(* IEC 61131-3 sources: plcassist-cli/packages/volt-lsp-iec/test-corpus/lenze-mid/Device/Plc Logic/Application/Library Manager/(unresolved)/visuusermgmt3 interfaces, 17 files *)

(* ---- VUM_CONSTANTS.gvl ---- *)
VAR_GLOBAL
	VISU_VUM_MAX_GROUPS_PER_USER : INT := 10;
END_VAR

(* ---- IEXTERNALUSERDATABASEPROVIDER.itf ---- *)
INTERFACE IEXTERNALUSERDATABASEPROVIDER
END_INTERFACE

METHOD CHANGEUSERPASSWORD : VUM_ReturnValues
VAR_INPUT
	WSTUSERNAME : WSTRING;
	WSTNEWPASSWORD : WSTRING;
	WSTOLDPASSWORD : WSTRING;
END_VAR
END_METHOD

METHOD CHECKLOGIN : VUM_ReturnValues
VAR_INPUT
	WSTUSERNAME : WSTRING;
	WSTPASSWORD : WSTRING;
END_VAR
VAR_OUTPUT
	WSTFULLNAME : WSTRING;
	DWUSERGROUPID : DWORD;
END_VAR
END_METHOD

METHOD CHECKLOGINWITHGROUPID : VUM_ReturnValues
VAR_INPUT
	WSTUSERNAME : WSTRING;
	WSTPASSWORD : WSTRING;
	DWUSERGROUPID : DWORD;
END_VAR
VAR_OUTPUT
	WSTFULLNAME : WSTRING;
END_VAR
END_METHOD

METHOD CHANGEUSER : VUM_ReturnValues
VAR_INPUT
	PVUMUSER : POINTER TO VUM_User;
	UDIINDEX : UDINT;
	EEDITTYPE : VUM_EditType;
END_VAR
END_METHOD

METHOD GETUSERCOUNT : UDINT
END_METHOD

METHOD GETUSERS : VUM_ReturnValues
VAR_INPUT
	UDISTARTINDEX : UDINT;
	UDIENDINDEX : UDINT;
	PARR : POINTER TO ARRAY [0..0] OF VUM_User;
	UDIARRSIZE : UDINT;
END_VAR
END_METHOD

(* ---- IEXTERNALUSERDATABASEPROVIDER2.itf ---- *)
INTERFACE IEXTERNALUSERDATABASEPROVIDER2
END_INTERFACE

METHOD FINDUSERBYTYPE : VUM_ReturnValues
VAR_INPUT
	VUMUSERIN : VUM_User;
	EEDITTYPE : VUM_EditType;
END_VAR
VAR_OUTPUT
	VUMUSER : VUM_User;
	UDIINDEX : UDINT;
END_VAR
END_METHOD

(* ---- IVISUUSERMANAGEMENT.itf ---- *)
INTERFACE IVISUUSERMANAGEMENT
END_INTERFACE

METHOD CHECKLOGIN : VUM_ReturnValues
VAR_INPUT
	WSTUSERNAME : WSTRING;
	WSTPASSWORD : WSTRING;
END_VAR
END_METHOD

METHOD CHECKLOGINWITHGROUPID : VUM_ReturnValues
VAR_INPUT
	WSTUSERNAME : WSTRING;
	WSTPASSWORD : WSTRING;
	DWUSERGROUPID : DWORD;
END_VAR
END_METHOD

METHOD REGISTEREXTERNALUSERDATABASEPROVIDER : VUM_ReturnValues
VAR_INPUT
	ITFEXTENALUSERDATABASEPROVIDER : IExternalUserDatabaseProvider;
END_VAR
END_METHOD

(* ---- IVISUUSERMANAGEMENT2.itf ---- *)
INTERFACE IVISUUSERMANAGEMENT2
END_INTERFACE

METHOD LOGINTOUSERGROUP : BOOL
VAR_INPUT
	PCLIENT : POINTER TO BYTE;
	DWGROUPID : DWORD;
	WSTUSERNAME : WSTRING(79);
	WSTFULLNAME : WSTRING(79);
END_VAR
END_METHOD

METHOD LOGINTOUSERGROUPS : BOOL
VAR_INPUT
	PCLIENT : POINTER TO BYTE;
	PADWUSERGROUPIDS : POINTER TO ARRAY [0..0] OF DWORD;
	DWUSERGROUPCOUNT : DWORD;
	WSTUSERNAME : WSTRING(79);
	WSTFULLNAME : WSTRING(79);
END_VAR
END_METHOD

(* ---- IVISUUSERMANAGEMENT3.itf ---- *)
INTERFACE IVISUUSERMANAGEMENT3
END_INTERFACE

METHOD CHANGEPASSWORD : VUM_ReturnValues
VAR_INPUT
	PCLIENT : POINTER TO BYTE;
	WSTUSERNAME : WSTRING(79);
	WSTNEWPASSWORD : WSTRING(79);
	WSTOLDPASSWORD : WSTRING(79);
END_VAR
END_METHOD

METHOD LOGIN : VUM_ReturnValues
VAR_INPUT
	PCLIENT : POINTER TO BYTE;
	WSTUSERNAME : WSTRING(79);
	WSTPASSWORD : WSTRING(79);
END_VAR
VAR_OUTPUT
	WSTFULLNAMEIFAVAILABLE : WSTRING;
	DWUSERGROUPID : DWORD;
	ADWUSERGROUPIDS : ARRAY [0..VUM_Constants.VISU_VUM_MAX_GROUPS_PER_USER] OF DWORD;
	DWUSERGROUPCOUNT : DWORD;
	BDEACTIVATED : BOOL;
END_VAR
END_METHOD

METHOD LOGOUT : VUM_ReturnValues
VAR_INPUT
	PCLIENT : POINTER TO BYTE;
END_VAR
END_METHOD

METHOD USERCOUNT : UDINT
VAR_INPUT
	PCLIENT : POINTER TO BYTE;
END_VAR
VAR_OUTPUT
	RESULT : VUM_ReturnValues;
END_VAR
END_METHOD

METHOD USERS : VUM_ReturnValues
VAR_INPUT
	PCLIENT : POINTER TO BYTE;
	UDISTARTINDEX : UDINT;
	UDIENDINDEX : UDINT;
	PARR : POINTER TO ARRAY [0..0] OF VUM_User2;
	UDIARRSIZE : UDINT;
END_VAR
END_METHOD

(* ---- IVISUUSERMANAGEMENT4.itf ---- *)
INTERFACE IVISUUSERMANAGEMENT4
END_INTERFACE

METHOD EDITUSER : VUM_ReturnValues
VAR_INPUT
	PCLIENT : POINTER TO BYTE;
	PVUMUSERNEW : POINTER TO VUM_User3;
	PVUMUSEROLD : POINTER TO VUM_User3;
	UDIINDEX : UDINT;
	EEDITTYPE : VUM_EditType;
END_VAR
END_METHOD

(* ---- IVISUUSERMGMTCHECKCHANGEUSERREQUESTPARAMETER.itf ---- *)
INTERFACE IVISUUSERMGMTCHECKCHANGEUSERREQUESTPARAMETER
END_INTERFACE

METHOD CHECKCHANGEUSERFLAGS : DWORD
END_METHOD

METHOD CHECKCHANGEUSERINDEX : DWORD
END_METHOD

METHOD CHECKCHANGEUSERTYPE : DWORD
END_METHOD

METHOD GETBUFFER : POINTER TO BYTE
VAR_INPUT
	XSWAPPINGNEEDED : BOOL;
END_VAR
END_METHOD

METHOD GETBUFFERSIZE : UDINT
END_METHOD

(* ---- IVISUUSERMGMTCHECKCHANGEUSERREQUESTRESULT.itf ---- *)
INTERFACE IVISUUSERMGMTCHECKCHANGEUSERREQUESTRESULT
END_INTERFACE

METHOD GETBUFFER : POINTER TO BYTE
END_METHOD

METHOD GETBUFFERSIZE : UDINT
END_METHOD

METHOD SETREADBYTES : BOOL
VAR_INPUT
	UDIREADBYTES : UDINT;
END_VAR
END_METHOD

METHOD SETRESULT
VAR_INPUT
	UDIRESULT : UDINT;
END_VAR
END_METHOD

(* ---- IVISUUSERMGMTCOMMONREQUESTPARAMETER.itf ---- *)
INTERFACE IVISUUSERMGMTCOMMONREQUESTPARAMETER
END_INTERFACE

METHOD GETREQUESTIDENTIFICATION : DataServerRequestIdentification
END_METHOD

METHOD GETREQUESTVERSION : DWORD
END_METHOD

METHOD GETUSERDB : DWORD
END_METHOD

(* ---- IVISUUSERMGMTCOMMONREQUESTRESULT.itf ---- *)
INTERFACE IVISUUSERMGMTCOMMONREQUESTRESULT
END_INTERFACE

METHOD SETERROR
VAR_INPUT
	UDIERROR : UDINT;
END_VAR
END_METHOD

METHOD SETRESULTVERSION
VAR_INPUT
	UDIVERSION : UDINT;
END_VAR
END_METHOD

METHOD SETSWAPPINGNEEDED
VAR_INPUT
	XSWAPPINGNEEDED : BOOL;
END_VAR
END_METHOD

(* ---- IVISUUSERMGMTGETSETDBREQUESTPARAMETER.itf ---- *)
INTERFACE IVISUUSERMGMTGETSETDBREQUESTPARAMETER
END_INTERFACE

METHOD GETSETDBFLAGS : DWORD
END_METHOD

(* ---- IVISUUSERMGMTGETSETDBREQUESTRESULT.itf ---- *)
INTERFACE IVISUUSERMGMTGETSETDBREQUESTRESULT
END_INTERFACE

METHOD SETUSERDB
VAR_INPUT
	UDIUSERDB : UDINT;
END_VAR
END_METHOD

(* ---- IVISUUSERMGMTGETUSERCOUNTREQUESTPARAMETER.itf ---- *)
INTERFACE IVISUUSERMGMTGETUSERCOUNTREQUESTPARAMETER
END_INTERFACE

(* ---- IVISUUSERMGMTGETUSERCOUNTREQUESTRESULT.itf ---- *)
INTERFACE IVISUUSERMGMTGETUSERCOUNTREQUESTRESULT
END_INTERFACE

METHOD SETUSERCOUNT
VAR_INPUT
	UDIUSERCOUNT : UDINT;
END_VAR
END_METHOD

(* ---- IVISUUSERMGMTGETUSERSREQUESTPARAMETER.itf ---- *)
INTERFACE IVISUUSERMGMTGETUSERSREQUESTPARAMETER
END_INTERFACE

METHOD GETENDINDEX : DWORD
END_METHOD

METHOD GETSTARTINDEX : DWORD
END_METHOD

(* ---- IVISUUSERMGMTGETUSERSREQUESTRESULT.itf ---- *)
INTERFACE IVISUUSERMGMTGETUSERSREQUESTRESULT
END_INTERFACE

METHOD GETBUFFER : POINTER TO BYTE
END_METHOD

METHOD GETBUFFERSIZE : UDINT
END_METHOD

METHOD SETREADBYTES : BOOL
VAR_INPUT
	UDIREADBYTES : UDINT;
END_VAR
END_METHOD
